Fanuc KAREL source: KO00104.KL

PROGRAM KO00104
%NOLOCKGROUP
VAR
  A: INTEGER
  B: ARRAY[2] OF SHORT
  OUT: REAL
BEGIN
  A = 1
  B[1] = 2
  OUT = ATAN2(A, B[1])
END KO00104
